// TIA Portal V20 export
// export: Created 2026-10-20T12:58:44.7433669Z, ExportSetting None, DisplayName Totally Integrated Automation Portal, DisplayVersion V20 Update 6, DisplayName TIA Portal Openness, DisplayVersion V20 Update 6, DisplayName TIA Portal Version Control Interface, DisplayVersion V20 Update 6, DisplayName SINAMICS Startdrive Advanced, DisplayVersion V20 SP1, DisplayName SINAMICS Startdrive G130, G150, S120, S150, SINAMICS MV, G220, S200, S210, DisplayVersion V20 SP1, DisplayName SINAMICS Startdrive G110M, G120, G120C, G120D, G120P, G115D, DisplayVersion V20 SP1, DisplayName STEP 7 Professional, DisplayVersion V20 Update 6, DisplayName STEP 7 Safety, DisplayVersion V20 Update 2, DisplayName WinCC Basic/Comfort/Advanced, DisplayVersion V20 Update 6, DisplayName WinCC Unified, DisplayVersion V20 Update 6
VAR_GLOBAL   // PLC tag table "Default tag table"
   RESET AT %I0.0 : Bool;
   "I-Device_Input_Main" AT %IW14 : Int;
   "I-Device_Output_Main" AT %QW14 : Int;
   Errors_Profinet_1 AT %MW8 : Word;
   HMI_Box_Connected_Main AT %MW10 : UInt;
   "I-Device_Input_System_1" AT %IW38 : Int;
   "I-Device_Output_System_1" AT %QW38 : Int;
   HMI_Box_Connected_2 AT %MW14 : UInt;
   HMI_Box_Connected_3 AT %MW16 : UInt;
   HMI_Box_Connected_5 AT %MW20 : UInt;
   HMI_Box_Connected_4 AT %MW18 : UInt;
   HMI_Box_Connected_1 AT %MW12 : UInt;
   "Profinet_HMI 1" AT %Q8.1 : Bool;
   "HMI 1 Estop" AT %Q8.0 : Bool;
   "Profinet_HMI 2" AT %Q8.3 : Bool;
   "HMI 2 Estop" AT %Q8.2 : Bool;
   System_Byte AT %MB1 : Byte;
   FirstScan AT %M1.0 : Bool;
   DiagStatusUpdate AT %M1.1 : Bool;
   AlwaysTRUE AT %M1.2 : Bool;
   AlwaysFALSE AT %M1.3 : Bool;
   Clock_Byte AT %MB0 : Byte;
   Clock_10Hz AT %M0.0 : Bool;
   Clock_5Hz AT %M0.1 : Bool;
   "Clock_2.5Hz" AT %M0.2 : Bool;
   Clock_2Hz AT %M0.3 : Bool;
   "Clock_1.25Hz" AT %M0.4 : Bool;
   Clock_1Hz AT %M0.5 : Bool;
   "Clock_0.625Hz" AT %M0.6 : Bool;
   "Clock_0.5Hz" AT %M0.7 : Bool;
   HMI_Communication_Lost AT %M6.0 : Bool;
   Heartbeat AT %MW2 : UInt;
   Heartbeat_ACK AT %MW4 : UInt;
   Reset_Comissioning AT %M10.1 : Bool;
   ACK AT %M10.0 : Bool;
   HMI_Reconnected AT %M10.3 : Bool;
   Error_Profinet_HMI_1 AT %M10.2 : Bool;
   Error_Profinet_HMI_2 AT %M10.4 : Bool;
END_VAR
